// TIA Portal V20 export
Screen "SYSTEM_SETTINGS_1"  1276x673
  ScreenItem "Title_ScreenOverview_X390_Y2" at 390,2 size 510x57  Type=HmiTextBox
  ScreenItem "Line_Header_X0_Y64" at 0,64 size 1280x0  Type=HmiLine
  ScreenItem "Frame_StandardProperties_1" at 825,327 size 350x121  Type=HmiRectangle
  ScreenItem "Frame_HMIData" at 825,70 size 350x121  Type=HmiRectangle
  ScreenItem "Frame_StandardProperties" at 465,70 size 350x121  Type=HmiRectangle
  ScreenItem "Frame_SafetyData" at 465,201 size 350x121  Type=HmiRectangle
  ScreenItem "Frame_PLC_Checksum" at 105,332 size 710x121  Type=HmiRectangle
  ScreenItem "Checksum_Textlists_DateTime" at 222,422 size 215x25  Type=HmiIOField
  ScreenItem "Text_Before" at 635,334 size 170x25  Type=HmiTextBox
  ScreenItem "Text_Safety_Checksum_1" at 107,395 size 110x25  Type=HmiTextBox
  ScreenItem "Checksum_Safety_Current" at 438,395 size 185x25  Type=HmiIOField
  ScreenItem "Checksum_Safety_Before" at 625,395 size 185x25  Type=HmiIOField
  ScreenItem "Text_Textlists_Checksum" at 107,422 size 110x25  Type=HmiTextBox
  ScreenItem "Checksum_Textlists_Current" at 438,422 size 185x25  Type=HmiIOField
  ScreenItem "Checksum_Textlists_Before" at 625,422 size 185x25  Type=HmiIOField
  ScreenItem "Text_DateTime" at 311,335 size 120x25  Type=HmiTextBox
  ScreenItem "Checksum_Standard_DateTime" at 222,368 size 215x25  Type=HmiIOField
  ScreenItem "Checksum_Safety_DateTime" at 222,395 size 215x25  Type=HmiIOField
  ScreenItem "Checksum_Standard_Before" at 625,368 size 185x25  Type=HmiIOField
  ScreenItem "Frame_Checksum_Standard_DateTime" at 221,367 size 217x27  Type=HmiRectangle
  ScreenItem "Frame_Checksum_Textlists_Current" at 437,421 size 187x27  Type=HmiRectangle
  ScreenItem "Frame_Checksum_Safety_DateTime" at 221,394 size 217x27  Type=HmiRectangle
  ScreenItem "Frame_Checksum_Standard_Current" at 437,367 size 187x27  Type=HmiRectangle
  ScreenItem "Title_PLC-Checksum" at 106,333 size 170x25  Type=HmiTextBox
  ScreenItem "Text_Current" at 453,334 size 170x25  Type=HmiTextBox
  ScreenItem "Text_Standard_Checksum" at 107,368 size 110x25  Type=HmiTextBox
  ScreenItem "Checksum_Standard_Current" at 438,368 size 185x25  Type=HmiIOField
  ScreenItem "Frame_Checksum_Textlists_DateTime" at 221,421 size 217x27  Type=HmiRectangle
  ScreenItem "Title_SMC-Diag" at 826,328 size 145x25  Type=HmiTextBox
  ScreenItem "Bar_SMCAssignedIn" at 1006,344 size 148x10  Type=HmiBar
  ScreenItem "Text_" at 1154,344 size 14x10  Type=HmiTextBox
  ScreenItem "IOField_WarningFromMemorySpace" at 954,390 size 50x25  Type=HmiIOField
  ScreenItem "IOField_AlarmFromMemorySpace" at 1118,390 size 50x25  Type=HmiIOField
  ScreenItem "Frame_Checksum_Safety_Current" at 437,394 size 187x27  Type=HmiRectangle
  ScreenItem "Rectangle_UsedLifetimeRed" at 953,416 size 52x27  Type=HmiRectangle
  ScreenItem "IOField_SMCAssigned" at 1083,362 size 85x25  Type=HmiIOField
  ScreenItem "IOField_SMCMemorySize" at 919,362 size 85x25  Type=HmiIOField
  ScreenItem "IOField_UsedLifetime" at 954,417 size 50x25  Type=HmiIOField
  ScreenItem "IOField_ParaLifetime" at 1118,417 size 50x25  Type=HmiIOField
  ScreenItem "Rectangle_SMCAssignedOrange" at 1082,362 size 87x27  Type=HmiRectangle
  ScreenItem "Rectangle_SMCAssignedRed" at 1082,362 size 87x27  Type=HmiRectangle
  ScreenItem "Text_ParaLifetime" at 1005,417 size 110x25  Type=HmiTextBox
  ScreenItem "PLCPropertiesMaxCycleTime" at 677,106 size 90x25  Type=HmiIOField
  ScreenItem "Text_PLCMinPropertiesCycleTime" at 467,133 size 250x25  Type=HmiTextBox
  ScreenItem "PLCPropertiesMinCycleTime" at 677,133 size 90x25  Type=HmiIOField
  ScreenItem "Text_PLCPropertiesComm" at 467,160 size 250x25  Type=HmiTextBox
  ScreenItem "PLCPropertiesComm" at 677,160 size 90x25  Type=HmiIOField
  ScreenItem "Title_PLC-Settings" at 466,71 size 300x25  Type=HmiTextBox
  ScreenItem "Title_HMIData" at 826,71 size 170x25  Type=HmiTextBox
  ScreenItem "Text_HMINumber" at 827,106 size 180x25  Type=HmiTextBox
  ScreenItem "HMINumber" at 1069,106 size 100x25  Type=HmiIOField
  ScreenItem "Text_SMCMemorySize" at 827,362 size 105x25  Type=HmiTextBox
  ScreenItem "Text_UsedLifetime" at 827,417 size 125x25  Type=HmiTextBox
  ScreenItem "Text_WarningFromMemorySpace" at 827,390 size 125x25  Type=HmiTextBox
  ScreenItem "Text_SMCAssigned" at 1005,362 size 90x25  Type=HmiTextBox
  ScreenItem "Text_AlarmFromMemorySpace" at 1005,390 size 110x25  Type=HmiTextBox
  ScreenItem "Text_PLCMaxPropertiesCycleTime" at 467,106 size 250x25  Type=HmiTextBox
  ScreenItem "Title_PLC-SafetyData_1" at 106,202 size 225x25  Type=HmiTextBox
  ScreenItem "Text_PLCSafetyMinCycleTime" at 107,264 size 240x25  Type=HmiTextBox
  ScreenItem "Text_PLCSafetyMaxCycleTime" at 107,291 size 240x25  Type=HmiTextBox
  ScreenItem "PLCSafatyMinCycleTime" at 350,264 size 90x25  Type=HmiIOField
  ScreenItem "PLCSafetyMaxCycleTime" at 350,291 size 90x25  Type=HmiIOField
  ScreenItem "Title_SafetyModeDeaktiv" at 636,204 size 225x25  Type=HmiTextBox
  ScreenItem "Text_FSignatur" at 467,237 size 150x25  Type=HmiTextBox
  ScreenItem "Title_PLC-SafetyData" at 466,203 size 160x25  Type=HmiTextBox
  ScreenItem "Text_FTimeStamp" at 467,264 size 150x25  Type=HmiTextBox
  ScreenItem "FTimeStamp" at 636,264 size 225x25  Type=HmiIOField
  ScreenItem "Title_SafetyModeAktiv" at 636,204 size 225x25  Type=HmiTextBox
  ScreenItem "FSignatur" at 636,237 size 225x25  Type=HmiIOField
  ScreenItem "PLCSafetyCycleTime" at 350,237 size 90x25  Type=HmiIOField
  ScreenItem "Text_PLCCycleTime" at 107,106 size 248x25  Type=HmiTextBox
  ScreenItem "PLCCycleTime" at 350,106 size 90x25  Type=HmiIOField
  ScreenItem "Title_PLC-StandardData" at 106,71 size 250x25  Type=HmiTextBox
  ScreenItem "Text_PLCMinCycleTime" at 107,133 size 248x25  Type=HmiTextBox
  ScreenItem "Text_PLCMaxCycleTime" at 107,160 size 248x25  Type=HmiTextBox
  ScreenItem "PLCMinCycleTime" at 350,133 size 90x25  Type=HmiIOField
  ScreenItem "PLCMaxCycleTime" at 350,160 size 90x25  Type=HmiIOField
  ScreenItem "Text_PLCSafetyCycleTime" at 107,237 size 240x25  Type=HmiTextBox
  ScreenItem "Title_PMLogon" at 827,133 size 100x25  Type=HmiTextBox
  ScreenItem "Text_CardUID" at 827,160 size 120x25  Type=HmiTextBox
  ScreenItem "Text_NoCard" at 1015,133 size 150x25  Type=HmiTextBox
  ScreenItem "Text_CardAvailable" at 1015,133 size 150x25  Type=HmiTextBox
  ScreenItem "IOField_CardUID" at 951,160 size 220x25  Type=HmiIOField
  ScreenItem "Button_CurveFCycleTimes" at 105,201 size 345x121  Type=HmiButton
  ScreenItem "Button_CurveStdCycleTimes" at 105,70 size 345x121  Type=HmiButton
  ScreenItem "Button_SICARHelp" at 1182,2 size 90x60  Type=HmiButton
  ScreenItem "Button_Language" at 1183,137 size 90x60  Type=HmiButton
  ScreenItem "Button_UpdateSMC" at 1183,204 size 90x60  Type=HmiButton
  ScreenItem "Button_DeleteBuffer" at 1090,2 size 90x60  Type=HmiButton
  ScreenItem "Button_Stop RT" at 1184,271 size 90x60  Type=HmiButton
  ScreenItem "Button_ResetFMinMaxTimes" at 1,201 size 90x60  Type=HmiButton
  ScreenItem "Button_ResetStdMinMaxTimes" at 1,70 size 90x60  Type=HmiButton
  ScreenItem "Button_SaveSettings" at 1183,70 size 90x60  Type=HmiButton
  ScreenItem "Button_SystemSettings" at 94,2 size 90x60  Type=HmiButton
  ScreenItem "Button_UpdateSMC_1" at 1,332 size 90x60  Type=HmiButton
  ScreenItem "permanentareaborderrectangle" at 0,0 size 0x0  Type=HmiRectangle
  ScreenItem "Button_Back" at 2,2 size 90x60  Type=HmiButton
